(* PLC project GeneratedProgram, SafePLC-Gen SafePLC-Gen Multimodal 1.0 *)
(* stored: creationDateTime 2026-04-25T14:00:19.203369Z *)

PROGRAM GeneratedProgram
  VAR
    TICSA_4750_03_Scaled : REAL;
    PICSA_4712_02_Scaled : REAL;
    PI_4712_01_Scaled : REAL;
    TICSA_4750_03_HH_SP : REAL;
    TICSA_4750_03_H_SP : REAL;
    TICSA_4750_03_L_SP : REAL;
    TICSA_4750_03_LL_SP : REAL;
    TICSA_4750_03_Deadband : REAL;
    PICSA_4712_02_HH_SP : REAL;
    PICSA_4712_02_H_SP : REAL;
    PICSA_4712_02_L_SP : REAL;
    PICSA_4712_02_LL_SP : REAL;
    PICSA_4712_02_Deadband : REAL;
    PI_4712_01_HH_SP : REAL;
    PI_4712_01_H_SP : REAL;
    PI_4712_01_L_SP : REAL;
    PI_4712_01_LL_SP : REAL;
    PI_4712_01_Deadband : REAL;
    TICSA_4750_03_HH : BOOL;
    TICSA_4750_03_H : BOOL;
    TICSA_4750_03_L : BOOL;
    TICSA_4750_03_LL : BOOL;
    TICSA_4750_03_HH_Ack : BOOL;
    TICSA_4750_03_LL_Ack : BOOL;
    TICSA_4750_03_HH_Set : BOOL;
    TICSA_4750_03_HH_Rst : BOOL;
    TICSA_4750_03_LL_Set : BOOL;
    TICSA_4750_03_LL_Rst : BOOL;
    TICSA_4750_03_HH_Latch : SR;
    TICSA_4750_03_LL_Latch : SR;
    PICSA_4712_02_HH : BOOL;
    PICSA_4712_02_H : BOOL;
    PICSA_4712_02_L : BOOL;
    PICSA_4712_02_LL : BOOL;
    PICSA_4712_02_HH_Ack : BOOL;
    PICSA_4712_02_LL_Ack : BOOL;
    PICSA_4712_02_HH_Set : BOOL;
    PICSA_4712_02_HH_Rst : BOOL;
    PICSA_4712_02_LL_Set : BOOL;
    PICSA_4712_02_LL_Rst : BOOL;
    PICSA_4712_02_HH_Latch : SR;
    PICSA_4712_02_LL_Latch : SR;
    PI_4712_01_HH : BOOL;
    PI_4712_01_H : BOOL;
    PI_4712_01_L : BOOL;
    PI_4712_01_LL : BOOL;
    PI_4712_01_HH_Ack : BOOL;
    PI_4712_01_LL_Ack : BOOL;
    PI_4712_01_HH_Set : BOOL;
    PI_4712_01_HH_Rst : BOOL;
    PI_4712_01_LL_Set : BOOL;
    PI_4712_01_LL_Rst : BOOL;
    PI_4712_01_HH_Latch : SR;
    PI_4712_01_LL_Latch : SR;
    LOOP_4750_03_TRIP : BOOL;
    LOOP_4712_02_TRIP : BOOL;
    SAFE_STATE : BOOL;
    TICSA_4750_03_SP : REAL;
    TICSA_4750_03_Error : REAL;
    TICSA_4750_03_Integral : REAL;
    TICSA_4750_03_Kp : REAL;
    TICSA_4750_03_Ki : REAL;
    TICSA_4750_03_Output : REAL;
    PICSA_4712_02_SP : REAL;
    PICSA_4712_02_Error : REAL;
    PICSA_4712_02_Integral : REAL;
    PICSA_4712_02_Kp : REAL;
    PICSA_4712_02_Ki : REAL;
    PICSA_4712_02_Output : REAL;
    FC_VALVE_Output : REAL;
    System_Alarm : BOOL;
    FirstScan : BOOL;
  END_VAR

            IF FirstScan THEN
    LOOP_4750_03_TRIP      := TRUE;
    LOOP_4712_02_TRIP      := TRUE;
    SAFE_STATE             := TRUE;
    TV_4750_03_Out         := 6554;
    PVA_4712_02_Out        := 6554;
    FC_VALVE_H_1007_IN_Out := 6554;
    SV_104_01              := FALSE;
    FirstScan              := FALSE;
    RETURN;
END_IF;

TICSA_4750_03_Scaled := ((INT_TO_REAL(TICSA_4750_03_Raw) - 6554.0) / (32767.0 - 6554.0)) * 150.0;
PICSA_4712_02_Scaled := ((INT_TO_REAL(PICSA_4712_02_Raw) - 6554.0) / (32767.0 - 6554.0)) * 10.0;
PI_4712_01_Scaled    := ((INT_TO_REAL(PI_4712_01_Raw)    - 6554.0) / (32767.0 - 6554.0)) * 10.0;

IF TICSA_4750_03_Scaled >= TICSA_4750_03_HH_SP THEN
    TICSA_4750_03_HH_Set := TRUE;
ELSIF TICSA_4750_03_Scaled <= (TICSA_4750_03_HH_SP - TICSA_4750_03_Deadband) THEN
    TICSA_4750_03_HH_Set := FALSE;
END_IF;
TICSA_4750_03_HH_Rst := TICSA_4750_03_HH_Ack AND (TICSA_4750_03_Scaled < TICSA_4750_03_HH_SP);
TICSA_4750_03_HH_Latch(S1 := TICSA_4750_03_HH_Set, R := TICSA_4750_03_HH_Rst);
TICSA_4750_03_HH := TICSA_4750_03_HH_Latch.Q1;

TICSA_4750_03_H := TICSA_4750_03_Scaled >= TICSA_4750_03_H_SP;
TICSA_4750_03_L := TICSA_4750_03_Scaled <= TICSA_4750_03_L_SP;

IF TICSA_4750_03_Scaled <= TICSA_4750_03_LL_SP THEN
    TICSA_4750_03_LL_Set := TRUE;
ELSIF TICSA_4750_03_Scaled >= (TICSA_4750_03_LL_SP + TICSA_4750_03_Deadband) THEN
    TICSA_4750_03_LL_Set := FALSE;
END_IF;
TICSA_4750_03_LL_Rst := TICSA_4750_03_LL_Ack AND (TICSA_4750_03_Scaled > TICSA_4750_03_LL_SP);
TICSA_4750_03_LL_Latch(S1 := TICSA_4750_03_LL_Set, R := TICSA_4750_03_LL_Rst);
TICSA_4750_03_LL := TICSA_4750_03_LL_Latch.Q1;

IF PICSA_4712_02_Scaled >= PICSA_4712_02_HH_SP THEN
    PICSA_4712_02_HH_Set := TRUE;
ELSIF PICSA_4712_02_Scaled <= (PICSA_4712_02_HH_SP - PICSA_4712_02_Deadband) THEN
    PICSA_4712_02_HH_Set := FALSE;
END_IF;
PICSA_4712_02_HH_Rst := PICSA_4712_02_HH_Ack AND (PICSA_4712_02_Scaled < PICSA_4712_02_HH_SP);
PICSA_4712_02_HH_Latch(S1 := PICSA_4712_02_HH_Set, R := PICSA_4712_02_HH_Rst);
PICSA_4712_02_HH := PICSA_4712_02_HH_Latch.Q1;

PICSA_4712_02_H := PICSA_4712_02_Scaled >= PICSA_4712_02_H_SP;
PICSA_4712_02_L := PICSA_4712_02_Scaled <= PICSA_4712_02_L_SP;

IF PICSA_4712_02_Scaled <= PICSA_4712_02_LL_SP THEN
    PICSA_4712_02_LL_Set := TRUE;
ELSIF PICSA_4712_02_Scaled >= (PICSA_4712_02_LL_SP + PICSA_4712_02_Deadband) THEN
    PICSA_4712_02_LL_Set := FALSE;
END_IF;
PICSA_4712_02_LL_Rst := PICSA_4712_02_LL_Ack AND (PICSA_4712_02_Scaled > PICSA_4712_02_LL_SP);
PICSA_4712_02_LL_Latch(S1 := PICSA_4712_02_LL_Set, R := PICSA_4712_02_LL_Rst);
PICSA_4712_02_LL := PICSA_4712_02_LL_Latch.Q1;

IF PI_4712_01_Scaled >= PI_4712_01_HH_SP THEN
    PI_4712_01_HH_Set := TRUE;
ELSIF PI_4712_01_Scaled <= (PI_4712_01_HH_SP - PI_4712_01_Deadband) THEN
    PI_4712_01_HH_Set := FALSE;
END_IF;
PI_4712_01_HH_Rst := PI_4712_01_HH_Ack AND (PI_4712_01_Scaled < PI_4712_01_HH_SP);
PI_4712_01_HH_Latch(S1 := PI_4712_01_HH_Set, R := PI_4712_01_HH_Rst);
PI_4712_01_HH := PI_4712_01_HH_Latch.Q1;

PI_4712_01_H := PI_4712_01_Scaled >= PI_4712_01_H_SP;
PI_4712_01_L := PI_4712_01_Scaled <= PI_4712_01_L_SP;

IF PI_4712_01_Scaled <= PI_4712_01_LL_SP THEN
    PI_4712_01_LL_Set := TRUE;
ELSIF PI_4712_01_Scaled >= (PI_4712_01_LL_SP + PI_4712_01_Deadband) THEN
    PI_4712_01_LL_Set := FALSE;
END_IF;
PI_4712_01_LL_Rst := PI_4712_01_LL_Ack AND (PI_4712_01_Scaled > PI_4712_01_LL_SP);
PI_4712_01_LL_Latch(S1 := PI_4712_01_LL_Set, R := PI_4712_01_LL_Rst);
PI_4712_01_LL := PI_4712_01_LL_Latch.Q1;

IF TICSA_4750_03_HH OR TICSA_4750_03_LL THEN
    LOOP_4750_03_TRIP := TRUE;
ELSIF LOOP_4750_03_TRIP AND MANUAL_RESET
      AND NOT TICSA_4750_03_HH AND NOT TICSA_4750_03_LL THEN
    LOOP_4750_03_TRIP := FALSE;
END_IF;

IF PICSA_4712_02_HH OR PICSA_4712_02_LL THEN
    LOOP_4712_02_TRIP := TRUE;
ELSIF LOOP_4712_02_TRIP AND MANUAL_RESET
      AND NOT PICSA_4712_02_HH AND NOT PICSA_4712_02_LL THEN
    LOOP_4712_02_TRIP := FALSE;
END_IF;

SAFE_STATE := ESTOP OR LOOP_4750_03_TRIP OR LOOP_4712_02_TRIP;

IF NOT SAFE_STATE THEN
    TICSA_4750_03_Error    := TICSA_4750_03_SP - TICSA_4750_03_Scaled;
    TICSA_4750_03_Integral := TICSA_4750_03_Integral + (TICSA_4750_03_Ki * TICSA_4750_03_Error);
    IF TICSA_4750_03_Integral > 100.0 THEN
        TICSA_4750_03_Integral := 100.0;
    ELSIF TICSA_4750_03_Integral < 0.0 THEN
        TICSA_4750_03_Integral := 0.0;
    END_IF;
    TICSA_4750_03_Output := (TICSA_4750_03_Kp * TICSA_4750_03_Error) + TICSA_4750_03_Integral;
    IF TICSA_4750_03_Output > 100.0 THEN
        TICSA_4750_03_Output := 100.0;
    ELSIF TICSA_4750_03_Output < 0.0 THEN
        TICSA_4750_03_Output := 0.0;
    END_IF;
    TV_4750_03_Out := REAL_TO_INT(6554.0 + (TICSA_4750_03_Output / 100.0) * (32767.0 - 6554.0));
ELSE
    TV_4750_03_Out := 6554;
END_IF;

IF NOT SAFE_STATE THEN
    PICSA_4712_02_Error    := PICSA_4712_02_SP - PICSA_4712_02_Scaled;
    PICSA_4712_02_Integral := PICSA_4712_02_Integral + (PICSA_4712_02_Ki * PICSA_4712_02_Error);
    IF PICSA_4712_02_Integral > 100.0 THEN
        PICSA_4712_02_Integral := 100.0;
    ELSIF PICSA_4712_02_Integral < 0.0 THEN
        PICSA_4712_02_Integral := 0.0;
    END_IF;
    PICSA_4712_02_Output := (PICSA_4712_02_Kp * PICSA_4712_02_Error) + PICSA_4712_02_Integral;
    IF PICSA_4712_02_Output > 100.0 THEN
        PICSA_4712_02_Output := 100.0;
    ELSIF PICSA_4712_02_Output < 0.0 THEN
        PICSA_4712_02_Output := 0.0;
    END_IF;
    PVA_4712_02_Out := REAL_TO_INT(6554.0 + (PICSA_4712_02_Output / 100.0) * (32767.0 - 6554.0));
ELSE
    PVA_4712_02_Out := 6554;
END_IF;

IF NOT SAFE_STATE THEN
    IF HS_4750_01 THEN
        FC_VALVE_Output := 100.0;
    ELSE
        FC_VALVE_Output := 0.0;
    END_IF;
    FC_VALVE_H_1007_IN_Out := REAL_TO_INT(6554.0 + (FC_VALVE_Output / 100.0) * (32767.0 - 6554.0));
ELSE
    FC_VALVE_H_1007_IN_Out := 6554;
END_IF;

SV_104_01 := NOT SAFE_STATE;

System_Alarm :=
    TICSA_4750_03_HH_Latch.Q1 OR TICSA_4750_03_LL_Latch.Q1 OR
    TICSA_4750_03_H            OR TICSA_4750_03_L            OR
    PICSA_4712_02_HH_Latch.Q1 OR PICSA_4712_02_LL_Latch.Q1 OR
    PICSA_4712_02_H            OR PICSA_4712_02_L            OR
    PI_4712_01_HH_Latch.Q1    OR PI_4712_01_LL_Latch.Q1    OR
    PI_4712_01_H               OR PI_4712_01_L              OR
    LOOP_4750_03_TRIP          OR LOOP_4712_02_TRIP         OR
    SAFE_STATE;
          
END_PROGRAM

CONFIGURATION Config0
  RESOURCE Res0 ON PLC
    TASK MainTask(INTERVAL := T#20ms, PRIORITY := 0);
    PROGRAM Main : GeneratedProgram;
  END_RESOURCE
END_CONFIGURATION
